(* IEC 61131-3 sources: bevling_machine/framework/sources, 2 files *)

(* ---- GVL_Motion.st ---- *)
(* 模块说明：旧单轴 Demo 的操作和监控变量。新切割机框架不使用这些变量；旧 Demo 当前未挂周期任务。 *)
VAR_GLOBAL
    (* 旧 Demo 操作命令：仅供单轴测试，新整机流程不使用。 *)
    xEnable     : BOOL; (* 旧 Demo 的 pandao 伺服使能请求，TRUE 上使能，FALSE 关闭。 *)
    xReset      : BOOL; (* 旧 Demo 轴故障复位请求，接 MC_Reset.Execute。 *)
    xStop       : BOOL; (* 旧 Demo 停止请求；停止完成后释放锁定，再决定是否重新启动。 *)
    xJogFwd     : BOOL; (* 历史正向点动入口，当前旧 Demo 正文未接入。 *)
    xJogRev     : BOOL; (* 历史反向点动入口，当前旧 Demo 正文未接入。 *)
    xMoveRel    : BOOL; (* 历史相对定位入口，当前旧 Demo 正文未接入。 *)
    xMoveAbs    : BOOL; (* 历史绝对定位入口，当前旧 Demo 正文未接入。 *)
    xStartCycle : BOOL; (* 旧 Demo 单次往返启动，上升沿有效；当前 Demo 未周期调用。 *)

    rRelDist    : LREAL := 100.0; (* 历史单次相对距离 mm，当前往返正文不采用该参数。 *)
    rTargetPos  : LREAL := 0.0; (* 历史绝对目标位置 mm，当前往返正文不采用该参数。 *)

    (* 旧 Demo 运动参数：实际采用及限幅见各参数同行说明。 *)
    rJogVel     : LREAL := 10.0; (* 历史点动速度 mm/s，当前往返正文不采用该参数。 *)
    rVel        : LREAL := 30.0; (* 旧 Demo 往返速度 mm/s，正文限幅为 1..10。 *)
    rAcc        : LREAL := 200.0; (* 旧 Demo 加速度 mm/s²，正文限幅为 10..200。 *)
    rDec        : LREAL := 200.0; (* 旧 Demo 减速度 mm/s²，正文限幅为 10..200。 *)
    rStroke     : LREAL := 100.0; (* 旧 Demo 请求的单程距离 mm，正文使用绝对值并限制最大 20。 *)
    tDwell      : TIME  := T#1S; (* 旧 Demo 每个行程端点停留时间。 *)

    (* 旧 Demo 运行反馈：仅在旧程序被调用时更新。 *)
    xPowered    : BOOL; (* MC_Power.Status，伺服已使能反馈。 *)
    xAxisReady  : BOOL; (* 旧 Demo 中由已使能、非忙、无错误组合得到的可用标志。 *)
    xBusy       : BOOL; (* 往返功能块或停止功能块正忙。 *)
    xDisabled   : BOOL; (* 旧 Demo 根据未使能得到的显示状态。 *)
    xStandStill : BOOL; (* 旧 Demo 根据已使能且非忙得到的显示状态，不是独立轴状态读取。 *)
    xStopping   : BOOL; (* 停止功能块正在执行。 *)
    xErrorStop  : BOOL; (* 旧 Demo 综合错误显示，与 xAxisError 同步。 *)
    xAxisError  : BOOL; (* 使能、往返、复位或停止功能块任一报错。 *)
    iAxisErrorID: DWORD; (* 历史错误码显示变量，当前正文未更新，需读取实际功能块 ErrorID。 *)
    rActPos     : LREAL; (* MC_ReadActualPosition 返回的 pandao 实际位置，单位 mm。 *)
    iState      : INT; (* 旧 Demo 当前 iCycle 步骤镜像，便于在线监控。 *)
END_VAR

(* ---- PLC_PRG.st ---- *)
(* 模块说明：周期入口：先解码实体面板，再解析通信、调度整机、发布反馈和映射逻辑输出，仅在 ETHERCAT1 调用一次。 *)
PROGRAM PLC_PRG
VAR
	fbPanel : FB_PanelInput; (* 实体/仿真面板解码实例，须先于通信和整机调度调用。 *)
	fbCommunication : FB_ModbusInterface; (* 通信命令解析和状态打包实例；打包的是上一扫描已发布的整机反馈。 *)
	fbMachine : FB_Machine; (* 整机调度实例，包含初始化、手动、自动、互锁、报警和设备管理。 *)
	fbIO : FB_IOMap; (* 逻辑 I/O 映射实例，当前只形成诊断需求，不驱动真实输出。 *)
	fbLamp : FB_Indicator; (* 面板两色指示灯逻辑实例；纯输出，不参与控制。 *)
	xSafetyBypassActive : BOOL; (* 安全许可两级旁路已生效；仅当一级开关与二级确认同时置位。 *)
END_VAR
PROGRAM PLC_PRG
(* 本程序只在 ETHERCAT1 中周期调用一次；内部功能块沿本调用链每扫描执行。 *)
(* 0. 面板物理点 -> 逻辑面板：常开/常闭等极性只在这层处理，接线接反改这里一行即可。
   用 xUseRealPanel 而不是 xSimulation 选来源，因为 xSimulation 必须恒为 TRUE（FALSE 整机报 3001），
   真实设备是靠 axRealDevice 逐台接管的，物理按钮与设备仿真必须能同时存在。 *)
IF GVL_Parameters.xUseRealPanel THEN
    GVL_IO.stPanelInputs.xAutoMode   := GVL_IO_Physical.xDiPanelAutoMode;
    GVL_IO.stPanelInputs.xInitialize := GVL_IO_Physical.xDiPanelInit;
    GVL_IO.stPanelInputs.xStart      := GVL_IO_Physical.xDiPanelStart;
    GVL_IO.stPanelInputs.xResetAlarm := GVL_IO_Physical.xDiPanelReset;
    GVL_IO.stPanelInputs.xRunStart   := GVL_IO_Physical.xDiPanelRunStart;
    (* 停止按钮是常闭触点：未按=TRUE、按下=FALSE。这里取反成"TRUE=按下"，
       物理下降沿在逻辑层变回上升沿，FB_Machine 只认一个沿，不用分两种按钮。 *)
    GVL_IO.stPanelInputs.xRunStop    := NOT GVL_IO_Physical.xDiPanelRunStop;
    (* 安全许可 = 旋钮在许可位 且 急停未按下。急停是常开触点，按下=TRUE=不安全。
       注意这是联锁逻辑，不是安全级回路；断线时读到 FALSE 会被当成"许可成立"。 *)
    GVL_IO.xSafetyOK := GVL_IO_Physical.xDiPanelSafetyPermit AND NOT GVL_IO_Physical.xDiEStop;
ELSE
    (* 仿真面板调试：许可沿用仿真设置，物理旋钮与急停不参与，否则没有面板时永远过不了许可。 *)
    GVL_IO.xSafetyOK := GVL_Simulation.stSettings.xSafetyOK;
END_IF
(* 先解码实体/仿真面板；模式旋钮为唯一模式来源，随后发布到只读监控接口。 *)
fbPanel(xSimulation:=GVL_Parameters.xSimulation,stReal:=GVL_IO.stPanelInputs,
    stSim:=GVL_Simulation.stPanelInputs,xContinuous:=GVL_Parameters.xContinuous,
    xUseRealPanel:=GVL_Parameters.xUseRealPanel);
GVL_Interface.stPanel:=fbPanel.stCommand;
(* 1. 解析上位机新命令并打包上一扫描状态，供本扫描整机处理。 *)
fbCommunication(xEnable:=GVL_Modbus.xEnable,stStatus:=GVL_Interface.stStatus,
    aStatus:=GVL_Interface.aDeviceStatus,awRx:=GVL_Modbus.awRx,awTx:=GVL_Modbus.awTx);
(* 2. 安全许可旁路：一级开关与二级确认同时置位才生效，单开关无效。
   旁路只替代安全许可旋钮，绝不能盖掉急停：急停按下时旁路同样失效。 *)
xSafetyBypassActive:=F_SafetyBypassActive(GVL_RealDevice.stSettings) AND NOT GVL_IO_Physical.xDiEStop;
(* 3. 整机选择操作来源，调度工序，通过互锁后统一调用设备。 *)
fbMachine(
	xSimulation:=GVL_Parameters.xSimulation,
	stPanel:=GVL_Interface.stPanel,
    stRemote:=fbCommunication.stCommand,
	xRemoteRequest:=fbCommunication.xRequest,
    xAllowRemoteStartStop:=GVL_Parameters.xAllowRemoteStartStop,
    wRemoteSequence:=fbCommunication.wRequestSequence,
	aManual:=GVL_Interface.aManual,
    stRecipe:=GVL_Parameters.stRecipe,
	stSim:=GVL_Simulation.stSettings,
    stReal:=GVL_RealDevice.stSettings,
	xSafetyBypassActive:=xSafetyBypassActive,
    xRealSafetyOK:=GVL_IO.xSafetyOK,
	xRealMaterial:=GVL_IO.xMaterialAtLength);
(* 4. 将整机反馈发布到监控接口，建议调试时从这里查看主步骤和支线步骤。 *)
GVL_Interface.stStatus:=fbMachine.stStatus;
GVL_Interface.aDeviceStatus:=fbMachine.aDeviceStatus;

(* 4.5 定长光电（设备 6）接管后，把它本扫描的到位状态发布成真实料信号。
    这里取的是刚算完的设备状态；FB_Machine 内部读的是上一扫描的同一个值，
    对送料这种等稳定信号的判断没有影响（扫描周期远小于去抖时间）。 *)
GVL_IO.xMaterialAtLength := fbMachine.aDeviceStatus[6].xActive;
(* 5. 形成逻辑输出并下沉到物理点；真实气缸阀电平在此写入 GVL_IO_Physical。 *)
fbIO(aCommand:=fbMachine.aSelectedCommand,
        aStatus:=fbMachine.aDeviceStatus,aValveOut:=fbMachine.aValveOut,aValveOutAux:=fbMachine.aValveOutAux,
        aG2Valve:=fbMachine.aG2Valve,uiG2Band:=fbMachine.uiG2Band,
    axOutputs:=GVL_IO.axDigitalOutputs);
(* 6. 面板指示灯：只读整机状态，不参与任何控制，放在最后算以保证与本扫描状态一致。 *)
fbLamp(xRunState:=fbMachine.stStatus.xRunState,eState:=fbMachine.stStatus.eState,
    eMode:=fbMachine.stStatus.eMode,udiAlarm:=fbMachine.stStatus.udiAlarm);
GVL_IO_Physical.xDoLampGreen:=fbLamp.xGreen;
GVL_IO_Physical.xDoLampRed:=fbLamp.xRed;
